(* IEC 61131-3 sources: teller/JD_Teller_LC2_V11/Network, 1 file *)

(* ---- ConfigObjects.st ---- *)
FUNCTION GLOBAL TAB TASK_CONF
_K_TASK, _K_REAL,
_K_END_VAR,

_K_TASK, _K_CYCLIC,
_K_END_VAR,

_K_TASK, _K_BACKGROUND,
_K_END_VAR,

_K_END_CONF
END_FUNCTION

FUNCTION GLOBAL TAB IPR_CONF
_K_IPR
	0$UINT,
_K_END_VAR,
_K_END_CONF
END_FUNCTION

FUNCTION GLOBAL TAB CONFIG_TABLES
00138$UINT,
0$UINT, 0, 7, "_ALARMDISPLAY",
0$UINT, 0, 4, "_ALARMX0PARA",
0$UINT, 0, 2, "_ALARMX1PARA",
0$UINT, 0, 2, "_ALARMX3PARA",
0$UINT, 0, 12, "_ALARMXBUFFER",
0$UINT, 0, 1, "_BIT32",
0$UINT, 0, 1, "_BIT32RAM",
0$UINT, 0, 3, "_CAN",
0$UINT, 1, 10, "_CANLIB",
0$UINT, 1, 14, "_FILESYS",
0$UINT, 2, 0, "_FIRSTALARM",
0$UINT, 0, 12, "_GLOBAL",
0$UINT, 0, 1, "_HOTALARM",
0$UINT, 0, 4, "_LANGUAGESELECTION",
0$UINT, 0, 1, "_LIMITMAX",
0$UINT, 0, 1, "_LIMITMIN",
0$UINT, 0, 95, "_LSE",
0$UINT, 1, 0, "_MULTITASK",
0$UINT, 0, 3, "_MYIO",
0$UINT, 0, 4, "_OSKERNEL",
0$UINT, 0, 6, "_OSZILSE",
0$UINT, 0, 0, "_OSZILSEBACKGROUND",
0$UINT, 0, 1, "_RADIO32",
0$UINT, 0, 1, "_RADIO32RAM",
0$UINT, 0, 2, "_SCREEN",
0$UINT, 0, 13, "_SCROLLAREA",
0$UINT, 0, 6, "_SCROLLAREA2",
0$UINT, 1, 31, "_SERLIB",
0$UINT, 0, 0, "_STDLIB",
0$UINT, 0, 5, "_SYSDATETIME",
0$UINT, 1, 1, "_TASKOBJECTCONTROL",
0$UINT, 0, 2, "_TOOLCAT",
0$UINT, 1, 10, "_VARANCANLIB",
0$UINT, 1, 10, "_VARANCANLIBOS",
0$UINT, 1, 20, "_VARANSERLIBOS",
0$UINT, 0, 1, "_XACCESS",
0$UINT, 0, 0, "ACTSCREENWINDOW",
0$UINT, 1, 20, "ASCII_BIN",
0$UINT, 1, 7, "BOX_EDITER",
0$UINT, 1, 6, "BOX_EDITOR_PREVIEW_TC",
0$UINT, 1, 0, "BOXGENERATOR",
0$UINT, 1, 23, "BUSINTERFACESDIASINTERNAL",
0$UINT, 2, 20, "CAICIOAINPUTCHANNEL",
0$UINT, 2, 20, "CAIINPUTCHANNEL",
0$UINT, 1, 0, "CALL_JAM_WINDOW",
0$UINT, 1, 50, "CDIAS2DATAMOVER",
0$UINT, 1, 0, "CHANNELBASEDATA",
0$UINT, 1, 0, "CHANNELBASEDATAWRITEONLY",
0$UINT, 2, 50, "CIO011_IM",
0$UINT, 2, 40, "CIO0XX",
0$UINT, 2, 20, "CIOOUTPUTCHANNEL",
0$UINT, 1, 61, "CIV521",
0$UINT, 2, 61, "CIV_BASE",
0$UINT, 5, 50, "CNC",
0$UINT, 0, 0, "CONTROLBYWRITE12_WRITEVALUE",
0$UINT, 1, 40, "CONTROLLER",
0$UINT, 0, 0, "COUNT_TO",
0$UINT, 2, 10, "DAIINPUTCHNL",
0$UINT, 1, 3, "DELAY_MACHINE",
0$UINT, 1, 50, "DIAS2DATAMOVER",
0$UINT, 2, 30, "DIASMASTER",
0$UINT, 1, 70, "DIASMASTERC",
0$UINT, 2, 10, "DIASMASTERMAIN",
0$UINT, 1, 0, "DIASMASTERPOSTSCAN",
0$UINT, 0, 0, "EASYFILEHANDLING",
0$UINT, 0, 0, "EASYFILELIST",
0$UINT, 1, 11, "EEPROM",
0$UINT, 0, 0, "ENCODER_INMETEN",
0$UINT, 1, 10, "ETV0551_IOS",
0$UINT, 1, 1, "ETV0555_IOS",
0$UINT, 1, 3, "ETVEDGE_DIGIO_BASE",
0$UINT, 0, 1, "FILE_IO",
0$UINT, 1, 0, "FILEBASE",
0$UINT, 1, 1, "FREE_JAMDETECTOR",
0$UINT, 0, 10, "GETBROADCASTDATA",
0$UINT, 0, 1, "GRAPHIC",
0$UINT, 1, 20, "HUB_BASE",
0$UINT, 2, 10, "HUB_BASE_ROOT",
0$UINT, 2, 30, "HWBASE",
0$UINT, 2, 50, "HWBASECDIAS",
0$UINT, 3, 0, "HWCONTROL",
0$UINT, 1, 10, "HWCONTROLBASE",
0$UINT, 1, 0, "HWRTPOSTSCAN",
0$UINT, 1, 6, "I2CCDIAS",
0$UINT, 1, 2, "INTERPOLATEXY_D",
0$UINT, 1, 0, "JAMDETECT_TELLER",
0$UINT, 1, 1, "JAMDETECTION_TEACHIN_TELLER",
0$UINT, 1, 0, "JD_OR_TELLER",
0$UINT, 1, 0, "LOADSAVEDATA",
0$UINT, 1, 5, "MACHINE_SETTINGS",
0$UINT, 1, 0, "MERKER",
0$UINT, 1, 18, "MERKEREX",
0$UINT, 1, 0, "OPERATORLOGIN_TELLER",
0$UINT, 1, 1, "PULSER",
0$UINT, 1, 3, "RAM",
0$UINT, 1, 16, "RAMEX",
0$UINT, 1, 8, "RAMFILE",
0$UINT, 1, 20, "REFERENCE",
0$UINT, 3, 0, "SAFETYCDIAS_BASE",
0$UINT, 1, 42, "SAFETYMANAGER",
0$UINT, 1, 3, "SCALE",
0$UINT, 1, 41, "SDIASBASE",
0$UINT, 1, 10, "SDIASHUBBASE",
0$UINT, 1, 57, "SDIASMANAGER",
0$UINT, 1, 26, "SDIASPLC",
0$UINT, 1, 0, "SERSEND",
0$UINT, 0, 0, "SETPASSWORD",
0$UINT, 0, 0, "SIGNAL_SPLITTER",
0$UINT, 1, 0, "SIGNAL_SPLITTER_BG_TELLER",
0$UINT, 1, 0, "SIMPULSJE_TELLER",
0$UINT, 1, 10, "STRING",
0$UINT, 1, 70, "STRINGINTERNAL",
0$UINT, 1, 10, "STRINGRAM",
0$UINT, 0, 0, "SUMMERTIME_SELECTOR",
0$UINT, 0, 0, "SV_HELP",
0$UINT, 1, 20, "SYNCCALL",
0$UINT, 0, 1, "SYSTEM",
0$UINT, 1, 0, "TANABECOUNTERSERIAL",
0$UINT, 1, 3, "TELLERCLASS_TELLER",
0$UINT, 0, 0, "TERMINALCONTROL",
0$UINT, 0, 0, "TIMECONVERT",
0$UINT, 1, 1, "TOOLCATHANDLING",
0$UINT, 1, 1, "TOOLLIGHT",
0$UINT, 2, 2, "VARAN_BASE",
0$UINT, 1, 40, "VARAN_CAN",
0$UINT, 1, 50, "VARAN_DATAMOVER",
0$UINT, 2, 12, "VARANMANAGER",
0$UINT, 1, 43, "VARANMANAGER_1",
0$UINT, 1, 20, "VARANMANAGER_BASE",
0$UINT, 1, 1, "VARANMANAGERPOSTSCAN",
0$UINT, 1, 3, "VIRTUALBASEINIT",
0$UINT, 1, 2, "VISU_BOXEDITER_MINMAX",
0$UINT, 0, 0, "VISU_JAM",
0$UINT, 1, 0, "VISUTELLER_TELLER",
0$UINT, 2, 10, "WATCHDOGDIAS",
0$UINT, 1, 0, "WISCOMMENT",
0$UINT, 0, 0, "WISFILTER",
0$UINT, 0, 0, "WRITE1",
ONE_CFG$UINT, 0, 0, "ONE_HardwareNet",
ONE_CFG$UINT, 0, 0, "ONE_JamDetection_Trombone",
ONE_CFG$UINT, 0, 0, "ONE_LseRtkAlarm",
ONE_CFG$UINT, 0, 0, "ONE_LseRtkMain",
ONE_CFG$UINT, 0, 0, "ONE_Teller",
ONE_CFG$UINT, 0, 0, "ONE_ToolCat",
TASK_CFG$UINT, 0, 0, "TASK_CONF",
IPR_CFG$UINT, 0, 0, "IPR_CONF",
PRJ_CFG$UINT, 0, 0, "JD_Teller_LC2_V11",
END_FUNCTION

#ifdef __LSLLDR_IOELEMENTS__
FUNCTION GLOBAL TAB _IO_ELEMENTS_TAB
0001$UINT, 0001$UINT,
"**IOCONN_EMPTY**", "CIO011_IM1.Encoder",
0020$UINT,
"**IOCONN_EMPTY**", "TellerClass1.iEncoder",
"**IOCONN_EMPTY**", "TellerClass1.iSensorSTR",
"**IOCONN_EMPTY**", "TellerClass1.iSensorL",
"**IOCONN_EMPTY**", "TellerClass1.iSensorR",
"**IOCONN_EMPTY**", "S11_Jamdetection_TeachIn_01.cSensor_03",
"**IOCONN_EMPTY**", "S11_Jamdetection_TeachIn_01.iEncoder",
"**IOCONN_EMPTY**", "TellerClass1.oHeadnr03",
"**IOCONN_EMPTY**", "TellerClass1.oHeadnr05",
"**IOCONN_EMPTY**", "TellerClass1.oHeadnr01",
"**IOCONN_EMPTY**", "TellerClass1.oHeadnr02",
"**IOCONN_EMPTY**", "JD_OR1.Out",
"**IOCONN_EMPTY**", "S11_Jamdetection_TeachIn_01.cSensor_01",
"**IOCONN_EMPTY**", "Encoder_Inmeten1.cEncoder",
"**IOCONN_EMPTY**", "S11_Jamdetection_TeachIn_01.cSensor_02",
"**IOCONN_EMPTY**", "SerSend1.Ser",
"**IOCONN_EMPTY**", "Read_serial1.RxTx",
"**IOCONN_EMPTY**", "JAMDETECT1.JamResetTanabe",
"**IOCONN_EMPTY**", "TellerClass1.oHeadnr04",
"**IOCONN_EMPTY**", "TellerClass1.cAnalogSpeedOut",
"**IOCONN_EMPTY**", "TellerClass1.cExtBoxCount",
END_FUNCTION
#endif //__LSLLDR_IOELEMENTS__

FUNCTION GLOBAL TAB CH_REDIRECT_EMB_TAB
0000$UINT,
00040$UINT,
"CIO011_IM;SerialNo", "\SerialNoStr.Data",
"CIO0xx;SerialNo", "\SerialNoStr.Data",
"CIV521;SerialNo", "\SerialNoStr.Data",
"HwBaseCDIAS;SerialNo", "\SerialNoStr.Data",
"OperatorLogIn_Teller;sOp01_Name", "\Op01_Name.Data",
"OperatorLogIn_Teller;sOp01_WW", "\Op01_WW.Data",
"OperatorLogIn_Teller;sOp02_Name", "\Op02_Name.Data",
"OperatorLogIn_Teller;sOp02_WW", "\Op02_WW.Data",
"OperatorLogIn_Teller;sOp03_Name", "\Op03_Name.Data",
"OperatorLogIn_Teller;sOp03_WW", "\Op03_WW.Data",
"OperatorLogIn_Teller;sOp04_Name", "\Op04_Name.Data",
"OperatorLogIn_Teller;sOp04_WW", "\Op04_WW.Data",
"OperatorLogIn_Teller;sOp05_Name", "\Op05_Name.Data",
"OperatorLogIn_Teller;sOp05_WW", "\Op05_WW.Data",
"OperatorLogIn_Teller;sOp06_Name", "\Op06_Name.Data",
"OperatorLogIn_Teller;sOp06_WW", "\Op06_WW.Data",
"OperatorLogIn_Teller;sOp07_Name", "\Op07_Name.Data",
"OperatorLogIn_Teller;sOp07_WW", "\Op07_WW.Data",
"OperatorLogIn_Teller;sOp08_Name", "\Op08_Name.Data",
"OperatorLogIn_Teller;sOp08_WW", "\Op08_WW.Data",
"OperatorLogIn_Teller;sOp09_Name", "\Op09_Name.Data",
"OperatorLogIn_Teller;sOp09_WW", "\Op09_WW.Data",
"OperatorLogIn_Teller;sOp10_Name", "\Op10_Name.Data",
"OperatorLogIn_Teller;sOp10_WW", "\Op10_WW.Data",
"OperatorLogIn_Teller;sOperator_Selected", "\Operator_Selected.Data",
"OperatorLogIn_Teller;sWW_Invoer", "\WW_Invoer.Data",
"SafetyCDIAS_Base;SerialNo", "\SerialNoStr.Data",
"SdiasBase;SerialNo", "\SerialNoStr.Data",
"ToolLight;BoxnameOutput", "\Boxname.Data",
"ToolLight;ExtFilter", "\FileHandling\ExtensionFilter.Data",
"ToolLight;toExtensionString", "\FileHandling\ExtensionFilter.Data",
"ToolLight;toFileString", "\FileHandling\FileString.Data",
"ToolLight;toPathString", "\FileHandling\PathString.Data",
"ToolLight;toSelFile", "\FileHandling\toOpenFileStr.Data",
"Varan_Base;SerialNo", "\SerialNoStr.Data",
"easyFileHandling;ExtensionFilterStr", "\ExtensionFilter.Data",
"easyFileHandling;FileStr", "\FileString.Data",
"easyFileHandling;PathStr", "\PathString.Data",
"easyFileHandling;toOpenFileSt", "\toOpenFileStr.Data",
"easyFileHandling;toOpenFileString", "\toOpenFileStr.Data",
END_FUNCTION
